FUNCTION_BLOCK FB_StandardConveyor EXTENDS FB_ConveyorBase

END_FUNCTION_BLOCK

(* stored: Version 1.1.0.1, ProductVersion 3.1 *)
